// // MIGRATION DRAFT: not included in PLC compilation.
// // Reference: Reference_Project/OPC_Control_FB.scl, object OPC_Control_FB.
// // Types, globals, calls, units and behavior require manual reconciliation.
// // See docs/TIA_Missing_Blocks.md before importing as PLC code.
FUNCTION_BLOCK OPC_Control_FB
// 
//    VAR_INPUT
//       Id : UInt;
//       All_In_Automatic : Bool;
//       VTD_Error : Bool;
//       OPC_Enable : Bool;
//       Clear_OrderTable : Bool;
//    END_VAR
// 
//    VAR_OUTPUT
//       Error_ID : Word;
//    END_VAR
// 
//    VAR
//       Source_Location   : ID_Decoded;
//       Destination_Location   : ID_Decoded;
//       State_Main : UInt;
//       State_VTD : UInt;
//       State_Shuttle : UInt;
//       State_CNV : UInt;
//       T_Wait_Report_Done   : TON;
//    END_VAR
// 
//    VAR_TEMP
//       i : UInt;
//       j : UInt;
//       f : UInt;
//       HMI_Reset : Bool;
//    END_VAR

// // MIGRATION DRAFT: not included in PLC compilation.
// // Reference: Reference_Project/OPC_Control_FB.scl, object OPC_Control_FB.
// // Types, globals, calls, units and behavior require manual reconciliation.
// // See docs/TIA_Missing_Blocks.md before importing as PLC code.
// IF FirstScan THEN
// 	    OPC_Enable := TRUE;
// 	END_IF;
// 
// 	    IF State_CNV > 0 AND State_CNV < 250 THEN
// 
// 	        IF Source_Location.Device_Type = 10 OR Destination_Location.Device_Type = 10 THEN
// 	            IF Control.LCnv_Sys[Id].Cnv_Level[Source_Location.Level].Cnv1.Error
// 	                OR
// 	                Control.LCnv_Sys[Id].Cnv_Level[Destination_Location.Level].Cnv1.Error THEN
// 	                Error_ID.%X3 := TRUE;
// 	                State_CNV := 400;
// 	            END_IF;
// 	        END_IF;
// 
// 	        IF Source_Location.Device_Type = 11 OR Destination_Location.Device_Type = 11 THEN
// 	            IF Control.LCnv_Sys[Id].Cnv_Level[Source_Location.Level].Cnv2.Error
// 	                OR
// 	                Control.LCnv_Sys[Id].Cnv_Level[Destination_Location.Level].Cnv2.Error THEN
// 	                Error_ID.%X3 := TRUE;
// 	                State_CNV := 400;
// 	            END_IF;
// 	        END_IF;
// 
// 	        IF Control.ECnv_Sys[Id].Error THEN
// 	            Error_ID.%X4 := TRUE;
// 	            State_CNV := 400;
// 	        END_IF;
// 	    END_IF;
// 
// 	    IF State_VTD > 0 AND State_VTD < 250 THEN
// 	        IF VTD_Error THEN
// 	            Error_ID.%X5 := TRUE;
// 	            State_VTD := 400;
// 	        END_IF;
// 	    END_IF;
// 
// 	    IF Reset_All THEN
// 	        Error_ID := 0;
// 	    END_IF;
// 
// 	IF State_VTD = 400 OR State_Shuttle = 400 OR State_CNV = 400 THEN
// 	    Error_ID.%X0 := TRUE;
// 	ELSE
// 	    Error_ID.%X0 := FALSE;
// 	    Error_ID.%X6 := FALSE;
// 	    Error_ID.%X7 := FALSE;
// 	    Error_ID.%X8 := FALSE;
// 	END_IF;
// 
// 	IF (Reset_All OR HMI_Reset) AND State_VTD = 400
// 	THEN
// 	    State_VTD := 250;
// 
// 	END_IF;
// 
// 	IF (Reset_All OR HMI_Reset) AND State_Shuttle = 400
// 	THEN
// 	    State_Shuttle := 250;
// 	END_IF;
// 
// 	IF (Reset_All OR HMI_Reset) AND State_CNV = 400
// 	THEN
// 	    State_CNV := 250;
// 	END_IF;
// 
// 	(*
// 	Type of task to be performed:
// 	    1 = Move to Floor
// 	    2 = Shuttle Transfer into VTD
// 	    3 = Shuttle Transfer out of VTD
// 	    4 = Transfer Pallet into VTD
// 	    5 = Transfer Pallet out of VTD
// 	    6 = Transfer Pallet Roller to Roller
// 	    7 = Transfer Pallet Chain to Chain
// 	    8 = Transfer to pick station
// 	    9 = Transfer from Pick station
// 	    10 = Weigh Pallet
// 	    11 = Set chain Cnv as active (lower)
// 	    12 = Set Roller Cnv as active (raise)
// 
// 	    Need to isolate ZZ in XXYYZZ to confirm i = ZZ
// 
// 	    Extract XX (first two digits)
// 	    xx := inputNumber / 10000;
// 
// 	    Extract YY (middle two digits)
// 	    yy := (inputNumber / 100) MOD 100;
// 
// 	    Extract ZZ (last two digits)
// 	    zz := inputNumber MOD 100;
// 	*)
// 
// 
// 	IF All_In_Automatic AND OPC_Enable THEN
// 
// 	        CASE State_Main OF
// 	            0:
// 	                State_Main := 10;
// 
// 	            10:
// 	                IF Control.WCS_OPC_Control[Id].Task_Data_Available AND
// 	                    State_VTD = 0 AND State_Shuttle = 0 AND State_CNV = 0 THEN
// 	                    State_Main := 20;
// 	                END_IF;
// 
// 	            20:
// 	                ID_Decode_F(ID := Control.WCS_OPC_Control[Id].Source_Location,
// 	                              ID_Decoded := Source_Location);
// 	                ID_Decode_F(ID := Control.WCS_OPC_Control[Id].Destination_Location,
// 	                              ID_Decoded := Destination_Location);
// 
// 
// 	                IF Control.WCS_OPC_Control[Id].Task_Type = 1
// 	                    AND NOT Control.VTD[Id].Running THEN
// 	                    State_VTD := 30;
// 	                    Control.WCS_OPC_Control[Id].Task_Data_Available := 0;
// 
// 
// 	                ELSIF Control.WCS_OPC_Control[Id].Task_Type = 2 OR Control.WCS_OPC_Control[Id].Task_Type = 3
// 	                THEN
// 	                    State_Shuttle := 70;
// 	                    Control.WCS_OPC_Control[Id].Task_Data_Available := 0;
// 
// 
// 	                ELSIF (Control.WCS_OPC_Control[Id].Task_Type = 4 OR Control.WCS_OPC_Control[Id].Task_Type = 5)
// 	                THEN
// 	                    State_CNV := 100;
// 	                    Control.WCS_OPC_Control[Id].Task_Data_Available := 0;
// 	                END_IF;
// 	        END_CASE;
// 
// 	            CASE State_VTD OF
// 	                0:
// 	                    ;
// 
// 	                30:
// 	                    State_Main := 0;
// 	                    Control.VTD[Id].Current_Task_Type := INT_TO_UINT(Control.WCS_OPC_Control[Id].Task_Type);
// 	                    Control.VTD[Id].Instruction.Pallet_Type := Control.WCS_OPC_Control[Id].Pallet_Type;
// 	                    Control.VTD[Id].Instruction.Task_ID := INT_TO_UINT(Control.WCS_OPC_Control[Id].Task_ID);
// 	                    Control.VTD[Id].Instruction.Task_Metadata := Control.WCS_OPC_Control[Id].Task_Metadata;
// 	                    Control.VTD[Id].Instruction.Move_To_Level := INT_TO_UINT(Destination_Location.Level);
// 	                    State_VTD := 35;
// 
// 
// 
// 
// 
// 
// 
// 
// 	                35:
// 	                    Control.WCS_OPC_Control[Id].SM_State := Control.VTD[Id].SM_State;
// 	                    IF Control.VTD[Id].Current_Level = Destination_Location.Level THEN
// 
// 	                        Control.WCS_OPC_Control[Id].Movement_Ready := TRUE;
// 	                        State_VTD := 41;
// 	                    ELSIF Control.VTD[Id].Enabled AND Control.VTD[Id].Running THEN
// 	                        Control.WCS_OPC_Control[Id].Movement_Ready := TRUE;
// 	                        State_VTD := 40;
// 	                    END_IF;
// 
// 	                40:
// 	                    Control.WCS_OPC_Control[Id].SM_State := Control.VTD[Id].SM_State;
// 	                    IF Control.VTD[Id].SM_State = 100 THEN
// 	                        State_VTD := 41;
// 	                    END_IF;
// 
// 	                41:
// 	                    T_Wait_Report_Done.TON(IN := TRUE,
// 	                                           PT := T#500ms);
// 	                   IF T_Wait_Report_Done.Q THEN
// 	                       Control.WCS_OPC_Control[Id].Movement_Request_Complete := TRUE;
// 	                       State_VTD := 45;
// 	                   END_IF;
// 
// 	                45:
// 	                    Control.WCS_OPC_Control[Id].SM_State := Control.VTD[Id].SM_State;
// 	                    IF Control.WCS_OPC_Control[Id].Movement_Request_Complete_Ack THEN
// 	                        State_VTD := 250;
// 	                    END_IF;
// 
// 	                250:
// 	                    Control.VTD[Id].Instruction.Reset := FALSE;
// 	                    Control.VTD[Id].Instruction.Pallet_Type := 0;
// 	                    Control.VTD[Id].Instruction.Task_ID := 0;
// 	                    Control.VTD[Id].Instruction.Task_Metadata := '';
// 	                    Control.VTD[Id].Instruction.Move_To_Level := 0;
// 	                    Control.VTD[Id].Current_Task_Type := 0;
// 
// 	                    IF (State_Shuttle = 0 OR State_Shuttle = 250) AND
// 	                        (State_CNV = 0 OR State_CNV = 250) THEN
// 
// 	                        Control.WCS_OPC_Control[Id].SM_State := 0;
// 	                        Control.WCS_OPC_Control[Id].Movement_Ready := FALSE;
// 	                        Control.WCS_OPC_Control[Id].Movement_Request_Complete := FALSE;
// 	                        Control.WCS_OPC_Control[Id].Movement_Request_Complete_Ack := FALSE;
// 	                        Control.WCS_OPC_Control[Id].Pallet_Weight := 0;
// 	                        Control.WCS_OPC_Control[Id].Task_Metadata := '';
// 	                        T_Wait_Report_Done.TON(IN := FALSE,
// 	                                               PT := T#0S);
// 	                       State_VTD := 0;
// 	                    END_IF;
// 
// 	                400:
// 	                    Error_ID.%X6 := TRUE;
// 	                    IF Reset_All OR HMI_Reset
// 	                    THEN
// 	                        Error_ID.%X5 := FALSE;
// 	                        Error_ID.%X6 := FALSE;
// 	                        State_VTD := 250;
// 	                    END_IF;
// 	            END_CASE;
// 	        END_REGION ;
// 
// 	            CASE State_Shuttle OF
// 	                0:
// 	                    ;
// 
// 	                70:
// 	                    State_Main := 0;
// 	                    Control.VTD[Id].Instruction.Task_ID := Control.WCS_OPC_Control[Id].Task_ID;
// 	                    Control.VTD[Id].Instruction.Task_Metadata := Control.WCS_OPC_Control[Id].Task_Metadata;
// 	                    Control.VTD[Id].Instruction.Pallet_Type := Control.WCS_OPC_Control[Id].Pallet_Type;
// 	                    Control.VTD[Id].Current_Task_Type := INT_TO_UINT(Control.WCS_OPC_Control[Id].Task_Type);
// 	                    Control.VTD[Id].Shuttle_Interlock.Shuttle_Interlock_Task_ID := INT_TO_UINT(Control.WCS_OPC_Control[Id].Task_ID);
// 	                    Control.VTD[Id].Shuttle_Interlock.Shuttle_Interlock_Task_Metadata := Control.WCS_OPC_Control[Id].Task_Metadata;
// 	                    Control.VTD[Id].Shuttle_Interlock.Shuttle_ID := INT_TO_UINT(Control.WCS_OPC_Control[Id].Shuttle_ID);
// 	                    Control.VTD[Id].Shuttle_Interlock.Shuttle_Loaded := Control.WCS_OPC_Control[Id].Shuttle_Loaded;
// 	                    Control.VTD[Id].Shuttle_Interlock.Shuttle_Start_Location := Control.WCS_OPC_Control[Id].Source_Location;
// 	                    Control.VTD[Id].Shuttle_Interlock.Shuttle_Target_Location := Control.WCS_OPC_Control[Id].Destination_Location;
// 
// 	                    Control.VTD[Id].Shuttle_Interlock.Interlock_Request := TRUE;
// 	                    State_Shuttle := 75;
// 
// 	                75:
// 	                    Control.WCS_OPC_Control[Id].SM_State := Control.VTD[Id].SM_State;
// 	                    IF Control.VTD[Id].Shuttle_Interlock.Ready_To_Interlock THEN
// 	                        Control.WCS_OPC_Control[Id].Movement_Ready := TRUE;
// 	                        Control.WCS_OPC_Control[Id].Task_Data_Available := FALSE;
// 	                        State_Shuttle := 80;
// 	                    END_IF;
// 
// 	                80:
// 	                    IF Control.VTD[Id].Shuttle_Interlock.Interlock_Complete THEN
// 	                        Control.VTD[Id].Shuttle_Interlock.Interlock_Request := FALSE;
// 	                        Control.WCS_OPC_Control[Id].Movement_Request_Complete := TRUE;
// 	                        State_Shuttle := 90;
// 	                    END_IF;
// 
// 
// 
// 
// 
// 
// 
// 
// 	                90:
// 	                    IF Control.WCS_OPC_Control[Id].Movement_Request_Complete_Ack THEN
// 	                        Control.VTD[Id].Shuttle_Interlock.Interlock_Complete_Ack := TRUE;
// 	                        State_Shuttle := 250;
// 	                    END_IF;
// 
// 	                250:
// 
// 	                    Control.VTD[Id].Shuttle_Interlock.Interlock_Request := FALSE;
// 	                    Control.VTD[Id].Shuttle_Interlock.Shuttle_Start_Location := 0;
// 	                    Control.VTD[Id].Shuttle_Interlock.Shuttle_Target_Location := 0;
// 	                    Control.VTD[Id].Shuttle_Interlock.Shuttle_Loaded := 0;
// 	                    Control.VTD[Id].Shuttle_Interlock.Shuttle_ID := 0;
// 	                    Control.VTD[Id].Shuttle_Interlock.Shuttle_Interlock_Task_ID := 0;
// 	                    Control.VTD[Id].Shuttle_Interlock.Shuttle_Interlock_Task_Metadata := '';
// 	                    Control.VTD[Id].Shuttle_Interlock.Interlock_Complete_Ack := FALSE;
// 
// 	                    IF (State_VTD = 0 OR State_VTD = 250) AND
// 	                        (State_CNV = 0 OR State_CNV = 250) THEN
// 
// 	                        Control.WCS_OPC_Control[Id].SM_State := 0;
// 	                        Control.WCS_OPC_Control[Id].Movement_Ready := FALSE;
// 	                        Control.WCS_OPC_Control[Id].Movement_Request_Complete := FALSE;
// 	                        Control.WCS_OPC_Control[Id].Movement_Request_Complete_Ack := FALSE;
// 	                        Control.WCS_OPC_Control[Id].Task_Metadata := '';
// 	                        T_Wait_Report_Done.TON(IN := FALSE,
// 	                                               PT := T#0S);
// 
// 	                        State_Shuttle := 0;
// 	                    END_IF;
// 
// 	                400:
// 	                    Error_ID.%X7 := TRUE;
// 	                    IF Reset_All OR HMI_Reset
// 	                    THEN
// 	                        Error_ID.%X7 := FALSE;
// 	                        State_Shuttle := 250;
// 	                    END_IF;
// 	            END_CASE;
// 	        END_REGION ;
// 
// 	            CASE State_CNV OF
// 	                0:
// 	                    ;
// 
// 	                100:
// 	                    State_Main := 0;
// 
// 
// 	                    IF Destination_Location.Level >= Settings_DB.VTD[Id].Lowest_Level AND Destination_Location.Level <= Settings_DB.VTD[Id].Highest_Level THEN
// 
// 
// 
// 	                        IF (Destination_Location.Device_Type = 10 AND Control.ECnv_Sys[Id].Cnv_Occupied AND
// 	                            NOT Control.LCnv_Sys[Id].Cnv_Level[Destination_Location.Level].Cnv1.Cnv_Occupied) OR
// 	                            (Destination_Location.Device_Type = 10 AND Destination_Location.Level = 1 AND Source_Location.Device_Type = 0 AND
// 	                            NOT Control.LCnv_Sys[Id].Cnv_Level[Destination_Location.Level].Cnv1.Cnv_Occupied)
// 	                        THEN
// 	                            Control.LCnv_Sys[Id].Cnv_Level[Destination_Location.Level].Cnv1.Instruction.Task_ID := INT_TO_UINT(Control.WCS_OPC_Control[Id].Task_ID);
// 	                            Control.LCnv_Sys[Id].Cnv_Level[Destination_Location.Level].Cnv1.Instruction.Task_Metadata := Control.WCS_OPC_Control[Id].Task_Metadata;
// 	                            Control.LCnv_Sys[Id].Cnv_Level[Destination_Location.Level].Cnv1.Current_Task_Type := INT_TO_UINT(Control.WCS_OPC_Control[Id].Task_Type);
// 	                            Control.LCnv_Sys[Id].Cnv_Level[Destination_Location.Level].Cnv1.Instruction.Transfer_From_ID := Control.WCS_OPC_Control[Id].Source_Location;
// 	                            Control.LCnv_Sys[Id].Cnv_Level[Destination_Location.Level].Cnv1.Instruction.Transfer_To_ID := Control.WCS_OPC_Control[Id].Destination_Location;
// 	                            IF Control.WCS_OPC_Control[Id].Pallet_Type = 'E' AND Control.WCS_OPC_Control[Id].Pallet_Alignment = 'L' THEN
// 	                                Control.LCnv_Sys[Id].Cnv_Level[Destination_Location.Level].Cnv1.Instruction.Pallet_Type := 3;
// 	                            ELSIF Control.WCS_OPC_Control[Id].Pallet_Type = 'E' AND Control.WCS_OPC_Control[Id].Pallet_Alignment = 'R' THEN
// 	                                Control.LCnv_Sys[Id].Cnv_Level[Destination_Location.Level].Cnv1.Instruction.Pallet_Type := 2;
// 	                            END_IF;
// 
// 
// 	                            Control.LCnv_Sys[Id].Cnv_Level[Destination_Location.Level].Cnv1.Instruction.Start_Transfer := TRUE;
// 	                            State_CNV := 105;
// 
// 
// 	                        ELSIF Destination_Location.Device_Type = 11 AND Control.ECnv_Sys[Id].Cnv_Occupied AND
// 	                            NOT Control.LCnv_Sys[Id].Cnv_Level[Destination_Location.Level].Cnv2.Cnv_Occupied
// 	                        THEN
// 	                            Control.LCnv_Sys[Id].Cnv_Level[Destination_Location.Level].Cnv2.Instruction.Task_ID := INT_TO_UINT(Control.WCS_OPC_Control[Id].Task_ID);
// 	                            Control.LCnv_Sys[Id].Cnv_Level[Destination_Location.Level].Cnv2.Instruction.Task_Metadata := Control.WCS_OPC_Control[Id].Task_Metadata;
// 	                            Control.LCnv_Sys[Id].Cnv_Level[Destination_Location.Level].Cnv2.Current_Task_Type := INT_TO_UINT(Control.WCS_OPC_Control[Id].Task_Type);
// 	                            Control.LCnv_Sys[Id].Cnv_Level[Destination_Location.Level].Cnv2.Instruction.Transfer_From_ID := Control.WCS_OPC_Control[Id].Source_Location;
// 	                            Control.LCnv_Sys[Id].Cnv_Level[Destination_Location.Level].Cnv2.Instruction.Transfer_To_ID := Control.WCS_OPC_Control[Id].Destination_Location;
// 	                            IF Control.WCS_OPC_Control[Id].Pallet_Type = 'E' AND Control.WCS_OPC_Control[Id].Pallet_Alignment = 'L' THEN
// 	                                Control.LCnv_Sys[Id].Cnv_Level[Destination_Location.Level].Cnv2.Instruction.Pallet_Type := 3;
// 	                            ELSIF Control.WCS_OPC_Control[Id].Pallet_Type = 'E' AND Control.WCS_OPC_Control[Id].Pallet_Alignment = 'R' THEN
// 	                                Control.LCnv_Sys[Id].Cnv_Level[Destination_Location.Level].Cnv2.Instruction.Pallet_Type := 2;
// 	                            END_IF;
// 
// 
// 	                            Control.LCnv_Sys[Id].Cnv_Level[Destination_Location.Level].Cnv2.Instruction.Start_Transfer := TRUE;
// 	                            State_CNV := 105;
// 
// 
// 	                        ELSIF (Destination_Location.Device_Type = 12 AND Source_Location.Device_Type = 10 AND
// 	                            NOT Control.ECnv_Sys[Id].Cnv_Occupied AND
// 	                            Control.LCnv_Sys[Id].Cnv_Level[Destination_Location.Level].Cnv1.Cnv_Occupied)
// 	                        THEN
// 	                            Control.ECnv_Sys[Id].Instruction.Task_ID := INT_TO_UINT(Control.WCS_OPC_Control[Id].Task_ID);
// 	                            Control.ECnv_Sys[Id].Instruction.Task_Metadata := Control.WCS_OPC_Control[Id].Task_Metadata;
// 	                            Control.ECnv_Sys[Id].Current_Task_Type := INT_TO_UINT(Control.WCS_OPC_Control[Id].Task_Type);
// 	                            Control.ECnv_Sys[Id].Instruction.Transfer_From_ID := Control.WCS_OPC_Control[Id].Source_Location;
// 	                            Control.ECnv_Sys[Id].Instruction.Transfer_To_ID := Control.WCS_OPC_Control[Id].Destination_Location;
// 	                            IF Control.WCS_OPC_Control[Id].Pallet_Type = 'E' AND Control.WCS_OPC_Control[Id].Pallet_Alignment = 'L' THEN
// 	                                Control.ECnv_Sys[Id].Instruction.Pallet_Type := 3;
// 	                            ELSIF Control.WCS_OPC_Control[Id].Pallet_Type = 'E' AND Control.WCS_OPC_Control[Id].Pallet_Alignment = 'R' THEN
// 	                                Control.ECnv_Sys[Id].Instruction.Pallet_Type := 2;
// 	                            ELSIF Control.WCS_OPC_Control[Id].Pallet_Type = 'E' AND Control.WCS_OPC_Control[Id].Pallet_Alignment = 'C' THEN
// 	                                Control.ECnv_Sys[Id].Instruction.Pallet_Type := 4;
// 	                            ELSIF Control.WCS_OPC_Control[Id].Pallet_Type = 'C' THEN
// 	                                Control.ECnv_Sys[Id].Instruction.Pallet_Type := 1;
// 	                            END_IF;
// 
// 
// 	                            Control.ECnv_Sys[Id].Instruction.Start_Transfer := TRUE;
// 	                            State_CNV := 105;
// 
// 
// 	                        ELSIF (Destination_Location.Device_Type = 12 AND Source_Location.Device_Type = 11 AND
// 	                            NOT Control.ECnv_Sys[Id].Cnv_Occupied AND
// 	                            Control.LCnv_Sys[Id].Cnv_Level[Destination_Location.Level].Cnv2.Cnv_Occupied)
// 	                        THEN
// 	                            Control.ECnv_Sys[Id].Instruction.Task_ID := INT_TO_UINT(Control.WCS_OPC_Control[Id].Task_ID);
// 	                            Control.ECnv_Sys[Id].Instruction.Task_Metadata := Control.WCS_OPC_Control[Id].Task_Metadata;
// 	                            Control.ECnv_Sys[Id].Current_Task_Type := INT_TO_UINT(Control.WCS_OPC_Control[Id].Task_Type);
// 	                            Control.ECnv_Sys[Id].Instruction.Transfer_From_ID := Control.WCS_OPC_Control[Id].Source_Location;
// 	                            Control.ECnv_Sys[Id].Instruction.Transfer_To_ID := Control.WCS_OPC_Control[Id].Destination_Location;
// 	                            IF Control.WCS_OPC_Control[Id].Pallet_Type = 'E' AND Control.WCS_OPC_Control[Id].Pallet_Alignment = 'L' THEN
// 	                                Control.ECnv_Sys[Id].Instruction.Pallet_Type := 3;
// 	                            ELSIF Control.WCS_OPC_Control[Id].Pallet_Type = 'E' AND Control.WCS_OPC_Control[Id].Pallet_Alignment = 'R' THEN
// 	                                Control.ECnv_Sys[Id].Instruction.Pallet_Type := 2;
// 	                            ELSIF Control.WCS_OPC_Control[Id].Pallet_Type = 'E' AND Control.WCS_OPC_Control[Id].Pallet_Alignment = 'C' THEN
// 	                                Control.ECnv_Sys[Id].Instruction.Pallet_Type := 4;
// 	                            ELSIF Control.WCS_OPC_Control[Id].Pallet_Type = 'C' THEN
// 	                                Control.ECnv_Sys[Id].Instruction.Pallet_Type := 1;
// 	                            END_IF;
// 
// 
// 	                            Control.ECnv_Sys[Id].Instruction.Start_Transfer := TRUE;
// 	                            State_CNV := 105;
// 
// 
// 	                        ELSIF (Destination_Location.Device_Type = Source_Location.Device_Type AND
// 	                            Control.LCnv_Sys[Id].Cnv_Level[Destination_Location.Level].Cnv1.Cnv_Occupied) AND
// 	                            Control.VTD[Id].Current_Level =  Settings_DB.LCnv_Sys[Id].Cnv_Level[Destination_Location.Level].Cnv1.Cnv_Level
// 	                        THEN
// 	                            Control.LCnv_Sys[Id].Cnv_Level[Destination_Location.Level].Cnv1.Instruction.Task_ID := INT_TO_UINT(Control.WCS_OPC_Control[Id].Task_ID);
// 	                            Control.LCnv_Sys[Id].Cnv_Level[Destination_Location.Level].Cnv1.Instruction.Task_Metadata := Control.WCS_OPC_Control[Id].Task_Metadata;
// 	                            Control.LCnv_Sys[Id].Cnv_Level[Destination_Location.Level].Cnv1.Current_Task_Type := INT_TO_UINT(Control.WCS_OPC_Control[Id].Task_Type);
// 	                            Control.LCnv_Sys[Id].Cnv_Level[Destination_Location.Level].Cnv1.Instruction.Transfer_From_ID := Control.WCS_OPC_Control[Id].Source_Location;
// 	                            Control.LCnv_Sys[Id].Cnv_Level[Destination_Location.Level].Cnv1.Instruction.Transfer_To_ID := Control.WCS_OPC_Control[Id].Destination_Location;
// 	                            IF Control.WCS_OPC_Control[Id].Pallet_Type = 'E' AND Control.WCS_OPC_Control[Id].Pallet_Alignment = 'L' THEN
// 	                                Control.LCnv_Sys[Id].Cnv_Level[Destination_Location.Level].Cnv1.Instruction.Pallet_Type := 3;
// 	                            ELSIF Control.WCS_OPC_Control[Id].Pallet_Type = 'E' AND Control.WCS_OPC_Control[Id].Pallet_Alignment = 'R' THEN
// 	                                Control.LCnv_Sys[Id].Cnv_Level[Destination_Location.Level].Cnv1.Instruction.Pallet_Type := 2;
// 	                            END_IF;
// 
// 
// 	                            Control.LCnv_Sys[Id].Cnv_Level[Destination_Location.Level].Cnv1.Instruction.Pallet_Allignment := TRUE;
// 	                            State_CNV := 112;
// 
// 
// 	                        ELSIF (Destination_Location.Device_Type = Source_Location.Device_Type AND
// 	                            Control.LCnv_Sys[Id].Cnv_Level[Destination_Location.Level].Cnv2.Cnv_Occupied) AND
// 	                            Control.VTD[Id].Current_Level =  Settings_DB.LCnv_Sys[Id].Cnv_Level[Destination_Location.Level].Cnv2.Cnv_Level
// 	                        THEN
// 	                            Control.LCnv_Sys[Id].Cnv_Level[Destination_Location.Level].Cnv2.Instruction.Task_ID := INT_TO_UINT(Control.WCS_OPC_Control[Id].Task_ID);
// 	                            Control.LCnv_Sys[Id].Cnv_Level[Destination_Location.Level].Cnv2.Instruction.Task_Metadata := Control.WCS_OPC_Control[Id].Task_Metadata;
// 	                            Control.LCnv_Sys[Id].Cnv_Level[Destination_Location.Level].Cnv2.Current_Task_Type := INT_TO_UINT(Control.WCS_OPC_Control[Id].Task_Type);
// 	                            Control.LCnv_Sys[Id].Cnv_Level[Destination_Location.Level].Cnv2.Instruction.Transfer_From_ID := Control.WCS_OPC_Control[Id].Source_Location;
// 	                            Control.LCnv_Sys[Id].Cnv_Level[Destination_Location.Level].Cnv2.Instruction.Transfer_To_ID := Control.WCS_OPC_Control[Id].Destination_Location;
// 	                            IF Control.WCS_OPC_Control[Id].Pallet_Type = 'E' AND Control.WCS_OPC_Control[Id].Pallet_Alignment = 'L' THEN
// 	                                Control.LCnv_Sys[Id].Cnv_Level[Destination_Location.Level].Cnv2.Instruction.Pallet_Type := 3;
// 	                            ELSIF Control.WCS_OPC_Control[Id].Pallet_Type = 'E' AND Control.WCS_OPC_Control[Id].Pallet_Alignment = 'R' THEN
// 	                                Control.LCnv_Sys[Id].Cnv_Level[Destination_Location.Level].Cnv2.Instruction.Pallet_Type := 2;
// 	                            END_IF;
// 
// 
// 	                            Control.LCnv_Sys[Id].Cnv_Level[Destination_Location.Level].Cnv2.Instruction.Pallet_Allignment := TRUE;
// 	                            State_CNV := 112;
// 	                        ELSE
// 	                            IF Destination_Location.Device_Type = 10 AND Control.LCnv_Sys[Id].Cnv_Level[Destination_Location.Level].Cnv1.Cnv_Occupied THEN
// 
// 	                                Control.LCnv_Sys[Id].Cnv_Level[Destination_Location.Level].Cnv1.Cnv_Errors.Error_Word_1.%X1 := TRUE;
// 
// 	                            ELSIF Destination_Location.Device_Type = 10 AND Control.LCnv_Sys[Id].Cnv_Level[Destination_Location.Level].Cnv1.Inputs.Shuttle_High THEN
// 
// 	                                Control.LCnv_Sys[Id].Cnv_Level[Destination_Location.Level].Cnv1.Cnv_Errors.Error_Word_1.%X2 := TRUE;
// 
// 	                            ELSIF Destination_Location.Device_Type = 11 AND Control.LCnv_Sys[Id].Cnv_Level[Destination_Location.Level].Cnv2.Cnv_Occupied THEN
// 
// 	                                Control.LCnv_Sys[Id].Cnv_Level[Destination_Location.Level].Cnv2.Cnv_Errors.Error_Word_1.%X1 := TRUE;
// 
// 	                            ELSIF Destination_Location.Device_Type = 11 AND Control.LCnv_Sys[Id].Cnv_Level[Destination_Location.Level].Cnv2.Inputs.Shuttle_High THEN
// 
// 	                                Control.LCnv_Sys[Id].Cnv_Level[Destination_Location.Level].Cnv2.Cnv_Errors.Error_Word_1.%X2 := TRUE;
// 
// 	                            ELSIF Destination_Location.Device_Type = 12 THEN
// 	                                Control.ECnv_Sys[Id].Cnv_Errors.Error_Word_1.%X1 := TRUE;
// 	                            END_IF;
// 
// 	                            State_CNV := 400;
// 	                        END_IF;
// 	                    END_IF;
// 
// 	                105:
// 
// 
// 	                    IF Source_Location.Level >= Settings_DB.VTD[Id].Lowest_Level AND Source_Location.Level <= Settings_DB.VTD[Id].Highest_Level THEN
// 
// 	                        IF Source_Location.Device_Type = 10 AND NOT Control.ECnv_Sys[Id].Cnv_Occupied AND
// 	                            Control.LCnv_Sys[Id].Cnv_Level[Source_Location.Level].Cnv1.Cnv_Occupied
// 	                        THEN
// 	                            Control.LCnv_Sys[Id].Cnv_Level[Source_Location.Level].Cnv1.Instruction.Task_ID := INT_TO_UINT(Control.WCS_OPC_Control[Id].Task_ID);
// 	                            Control.LCnv_Sys[Id].Cnv_Level[Source_Location.Level].Cnv1.Instruction.Task_Metadata := Control.WCS_OPC_Control[Id].Task_Metadata;
// 	                            Control.LCnv_Sys[Id].Cnv_Level[Source_Location.Level].Cnv1.Current_Task_Type := INT_TO_UINT(Control.WCS_OPC_Control[Id].Task_Type);
// 	                            Control.LCnv_Sys[Id].Cnv_Level[Source_Location.Level].Cnv1.Instruction.Transfer_To_ID := Control.WCS_OPC_Control[Id].Destination_Location;
// 	                            Control.LCnv_Sys[Id].Cnv_Level[Source_Location.Level].Cnv1.Instruction.Transfer_From_ID := Control.WCS_OPC_Control[Id].Source_Location;
// 
// 
// 	                            Control.LCnv_Sys[Id].Cnv_Level[Source_Location.Level].Cnv1.Instruction.Start_Transfer := TRUE;
// 	                            State_CNV := 110;
// 
// 
// 	                        ELSIF (Source_Location.Device_Type = 11 AND NOT Control.ECnv_Sys[Id].Cnv_Occupied AND
// 	                            Control.LCnv_Sys[Id].Cnv_Level[Source_Location.Level].Cnv2.Cnv_Occupied) OR
// 	                            (Source_Location.Device_Type = 11 AND Source_Location.Level = 1 AND Destination_Location.Device_Type = 0 AND
// 	                            Control.LCnv_Sys[Id].Cnv_Level[Destination_Location.Level].Cnv2.Cnv_Occupied)
// 	                        THEN
// 	                            Control.LCnv_Sys[Id].Cnv_Level[Source_Location.Level].Cnv2.Instruction.Task_ID := INT_TO_UINT(Control.WCS_OPC_Control[Id].Task_ID);
// 	                            Control.LCnv_Sys[Id].Cnv_Level[Source_Location.Level].Cnv2.Instruction.Task_Metadata := Control.WCS_OPC_Control[Id].Task_Metadata;
// 	                            Control.LCnv_Sys[Id].Cnv_Level[Source_Location.Level].Cnv2.Current_Task_Type := INT_TO_UINT(Control.WCS_OPC_Control[Id].Task_Type);
// 	                            Control.LCnv_Sys[Id].Cnv_Level[Source_Location.Level].Cnv2.Instruction.Transfer_To_ID := Control.WCS_OPC_Control[Id].Destination_Location;
// 	                            Control.LCnv_Sys[Id].Cnv_Level[Source_Location.Level].Cnv2.Instruction.Transfer_From_ID := Control.WCS_OPC_Control[Id].Source_Location;
// 
// 
// 	                            Control.LCnv_Sys[Id].Cnv_Level[Source_Location.Level].Cnv2.Instruction.Start_Transfer := TRUE;
// 	                            State_CNV := 110;
// 
// 
// 	                        ELSIF (Source_Location.Device_Type = 12 AND Destination_Location.Device_Type = 10 AND Control.ECnv_Sys[Id].Cnv_Occupied AND
// 	                            NOT Control.LCnv_Sys[Id].Cnv_Level[Source_Location.Level].Cnv1.Cnv_Occupied)
// 	                        THEN
// 	                            Control.ECnv_Sys[Id].Instruction.Task_ID := INT_TO_UINT(Control.WCS_OPC_Control[Id].Task_ID);
// 	                            Control.ECnv_Sys[Id].Instruction.Task_Metadata := Control.WCS_OPC_Control[Id].Task_Metadata;
// 	                            Control.ECnv_Sys[Id].Current_Task_Type := INT_TO_UINT(Control.WCS_OPC_Control[Id].Task_Type);
// 	                            Control.ECnv_Sys[Id].Instruction.Transfer_To_ID := Control.WCS_OPC_Control[Id].Destination_Location;
// 	                            Control.ECnv_Sys[Id].Instruction.Transfer_From_ID := Control.WCS_OPC_Control[Id].Source_Location;
// 
// 
// 	                            Control.ECnv_Sys[Id].Instruction.Start_Transfer := TRUE;
// 	                            State_CNV := 110;
// 
// 
// 	                        ELSIF (Source_Location.Device_Type = 12 AND Destination_Location.Device_Type = 11 AND Control.ECnv_Sys[Id].Cnv_Occupied AND
// 	                            NOT Control.LCnv_Sys[Id].Cnv_Level[Source_Location.Level].Cnv2.Cnv_Occupied)
// 	                        THEN
// 	                            Control.ECnv_Sys[Id].Instruction.Task_ID := INT_TO_UINT(Control.WCS_OPC_Control[Id].Task_ID);
// 	                            Control.ECnv_Sys[Id].Instruction.Task_Metadata := Control.WCS_OPC_Control[Id].Task_Metadata;
// 	                            Control.ECnv_Sys[Id].Current_Task_Type := INT_TO_UINT(Control.WCS_OPC_Control[Id].Task_Type);
// 	                            Control.ECnv_Sys[Id].Instruction.Transfer_To_ID := Control.WCS_OPC_Control[Id].Destination_Location;
// 	                            Control.ECnv_Sys[Id].Instruction.Transfer_From_ID := Control.WCS_OPC_Control[Id].Source_Location;
// 
// 
// 	                            Control.ECnv_Sys[Id].Instruction.Start_Transfer := TRUE;
// 	                            State_CNV := 110;
// 	                        ELSE
// 	                            State_CNV := 400;
// 	                        END_IF;
// 	                    ELSE
// 	                        State_CNV := 400;
// 	                    END_IF;
// 
// 	                110:
// 	                    Control.WCS_OPC_Control[Id].SM_State := Control.ECnv_Sys[Id].SM_State;
// 
// 	                    IF Control.ECnv_Sys[Id].Enabled AND Control.ECnv_Sys[Id].Running
// 	                    THEN
// 	                        Control.ECnv_Sys[Id].Instruction.Start_Transfer := FALSE;
// 	                        IF (Source_Location.Device_Type = 12 AND Destination_Location.Device_Type = 10) OR
// 	                            (Source_Location.Device_Type = 10 AND Destination_Location.Device_Type = 12) AND
// 	                            Control.LCnv_Sys[Id].Cnv_Level[Control.VTD[Id].Current_Level].Cnv1.Running
// 	                        THEN
// 	                            Control.LCnv_Sys[Id].Cnv_Level[Control.VTD[Id].Current_Level].Cnv1.Instruction.Start_Transfer := FALSE;
// 	                            State_CNV := 115;
// 	                        ELSIF (Source_Location.Device_Type = 12 AND Destination_Location.Device_Type = 11) OR
// 	                            (Source_Location.Device_Type = 11 AND Destination_Location.Device_Type = 12) AND
// 	                            Control.LCnv_Sys[Id].Cnv_Level[Control.VTD[Id].Current_Level].Cnv2.Running
// 	                        THEN
// 	                            Control.LCnv_Sys[Id].Cnv_Level[Control.VTD[Id].Current_Level].Cnv2.Instruction.Start_Transfer := FALSE;
// 	                            State_CNV := 115;
// 	                        END_IF;
// 	                        Control.WCS_OPC_Control[Id].Movement_Ready := TRUE;
// 	                    END_IF;
// 
// 	                112:
// 	                    IF Control.LCnv_Sys[Id].Cnv_Level[Destination_Location.Level].Cnv1.Enabled AND Control.LCnv_Sys[Id].Cnv_Level[Destination_Location.Level].Cnv1.Running
// 	                    THEN
// 	                        Control.WCS_OPC_Control[Id].SM_State := Control.LCnv_Sys[Id].Cnv_Level[Destination_Location.Level].Cnv1.SM_State;
// 	                        Control.LCnv_Sys[Id].Cnv_Level[Destination_Location.Level].Cnv1.Instruction.Pallet_Allignment := FALSE;
// 	                        Control.WCS_OPC_Control[Id].Movement_Ready := TRUE;
// 	                        State_CNV := 116;
// 	                    ELSIF Control.LCnv_Sys[Id].Cnv_Level[Destination_Location.Level].Cnv2.Enabled AND Control.LCnv_Sys[Id].Cnv_Level[Destination_Location.Level].Cnv2.Running
// 	                    THEN
// 	                        Control.WCS_OPC_Control[Id].SM_State := Control.LCnv_Sys[Id].Cnv_Level[Destination_Location.Level].Cnv2.SM_State;
// 	                        Control.LCnv_Sys[Id].Cnv_Level[Destination_Location.Level].Cnv2.Instruction.Pallet_Allignment := FALSE;
// 	                        Control.WCS_OPC_Control[Id].Movement_Ready := TRUE;
// 	                        State_CNV := 116;
// 	                    END_IF;
// 
// 
// 
// 	                115:
// 	                    Control.WCS_OPC_Control[Id].SM_State := Control.ECnv_Sys[Id].SM_State;
// 	                    IF (Source_Location.Device_Type = 12 AND Destination_Location.Device_Type = 10) OR
// 	                        (Source_Location.Device_Type = 10 AND Destination_Location.Device_Type = 12) THEN
// 	                        IF Control.ECnv_Sys[Id].Done AND Control.LCnv_Sys[Id].Cnv_Level[Destination_Location.Level].Cnv1.Done THEN
// 	                            State_CNV := 118;
// 	                        END_IF;
// 	                    ELSIF (Source_Location.Device_Type = 12 AND Destination_Location.Device_Type = 11) OR
// 	                        (Source_Location.Device_Type = 11 AND Destination_Location.Device_Type = 12) THEN
// 	                        IF Control.ECnv_Sys[Id].Done AND Control.LCnv_Sys[Id].Cnv_Level[Destination_Location.Level].Cnv2.Done THEN
// 	                            State_CNV := 118;
// 	                        END_IF;
// 	                    END_IF;
// 
// 	                116:
// 	                        IF Control.LCnv_Sys[Id].Cnv_Level[Destination_Location.Level].Cnv1.Done THEN
// 	                            State_CNV := 118;
// 	                        END_IF;
// 	                        IF Control.LCnv_Sys[Id].Cnv_Level[Destination_Location.Level].Cnv2.Done THEN
// 	                            State_CNV := 118;
// 	                        END_IF;
// 
// 	                118:
// 	                    T_Wait_Report_Done.TON(IN := TRUE,
// 	                                           PT := T#500mS);
// 	                   IF T_Wait_Report_Done.Q THEN
// 	                        Control.WCS_OPC_Control[Id].Movement_Request_Complete := TRUE;
// 	                        State_CNV := 120;
// 	                    END_IF;
// 
// 	                120:
// 	                    Control.WCS_OPC_Control[Id].SM_State := Control.ECnv_Sys[Id].SM_State;
// 	                    IF Control.WCS_OPC_Control[Id].Movement_Request_Complete_Ack THEN
// 	                        State_CNV := 250;
// 	                    END_IF;
// 
// 	                250:
// 	                    Control.ECnv_Sys[Id].Instruction.Reset := FALSE;
// 	                    Control.ECnv_Sys[Id].Instruction.Start_Transfer := FALSE;
// 	                    Control.ECnv_Sys[Id].Instruction.Task_ID := 0;
// 	                    Control.ECnv_Sys[Id].Instruction.Task_Metadata := '';
// 	                    Control.ECnv_Sys[Id].Current_Task_Type := 0;
// 	                    Control.ECnv_Sys[Id].Instruction.Transfer_From_ID := 0;
// 	                    Control.ECnv_Sys[Id].Instruction.Transfer_To_ID := 0;
// 	                    IF Destination_Location.Device_Type = 10 THEN
// 	                        Control.LCnv_Sys[Id].Cnv_Level[Destination_Location.Level].Cnv1.Instruction.Reset := FALSE;
// 	                        Control.LCnv_Sys[Id].Cnv_Level[Destination_Location.Level].Cnv1.Instruction.Start_Transfer := FALSE;
// 	                        Control.LCnv_Sys[Id].Cnv_Level[Destination_Location.Level].Cnv1.Instruction.Task_ID := 0;
// 	                        Control.LCnv_Sys[Id].Cnv_Level[Destination_Location.Level].Cnv1.Instruction.Task_Metadata := '';
// 	                        Control.LCnv_Sys[Id].Cnv_Level[Destination_Location.Level].Cnv1.Current_Task_Type := 0;
// 	                        Control.LCnv_Sys[Id].Cnv_Level[Destination_Location.Level].Cnv1.Instruction.Transfer_From_ID := 0;
// 	                        Control.LCnv_Sys[Id].Cnv_Level[Destination_Location.Level].Cnv1.Instruction.Transfer_To_ID := 0;
// 	                    ELSIF Destination_Location.Device_Type = 11 THEN
// 	                        Control.LCnv_Sys[Id].Cnv_Level[Destination_Location.Level].Cnv2.Instruction.Reset := FALSE;
// 	                        Control.LCnv_Sys[Id].Cnv_Level[Destination_Location.Level].Cnv2.Instruction.Start_Transfer := FALSE;
// 	                        Control.LCnv_Sys[Id].Cnv_Level[Destination_Location.Level].Cnv2.Instruction.Task_ID := 0;
// 	                        Control.LCnv_Sys[Id].Cnv_Level[Destination_Location.Level].Cnv2.Instruction.Task_Metadata := '';
// 	                        Control.LCnv_Sys[Id].Cnv_Level[Destination_Location.Level].Cnv2.Current_Task_Type := 0;
// 	                        Control.LCnv_Sys[Id].Cnv_Level[Destination_Location.Level].Cnv2.Instruction.Transfer_From_ID := 0;
// 	                        Control.LCnv_Sys[Id].Cnv_Level[Destination_Location.Level].Cnv2.Instruction.Transfer_To_ID := 0;
// 	                    ELSIF Source_Location.Device_Type = 10 THEN
// 	                        Control.LCnv_Sys[Id].Cnv_Level[Source_Location.Level].Cnv1.Instruction.Reset := FALSE;
// 	                        Control.LCnv_Sys[Id].Cnv_Level[Source_Location.Level].Cnv1.Instruction.Start_Transfer := FALSE;
// 	                        Control.LCnv_Sys[Id].Cnv_Level[Source_Location.Level].Cnv1.Instruction.Task_ID := 0;
// 	                        Control.LCnv_Sys[Id].Cnv_Level[Source_Location.Level].Cnv1.Instruction.Task_Metadata := '';
// 	                        Control.LCnv_Sys[Id].Cnv_Level[Source_Location.Level].Cnv1.Current_Task_Type := 0;
// 	                        Control.LCnv_Sys[Id].Cnv_Level[Source_Location.Level].Cnv1.Instruction.Transfer_From_ID := 0;
// 	                        Control.LCnv_Sys[Id].Cnv_Level[Source_Location.Level].Cnv1.Instruction.Transfer_To_ID := 0;
// 	                    ELSIF Destination_Location.Device_Type = 11 THEN
// 	                        Control.LCnv_Sys[Id].Cnv_Level[Source_Location.Level].Cnv2.Instruction.Reset := FALSE;
// 	                        Control.LCnv_Sys[Id].Cnv_Level[Source_Location.Level].Cnv2.Instruction.Start_Transfer := FALSE;
// 	                        Control.LCnv_Sys[Id].Cnv_Level[Source_Location.Level].Cnv2.Instruction.Task_ID := 0;
// 	                        Control.LCnv_Sys[Id].Cnv_Level[Source_Location.Level].Cnv2.Instruction.Task_Metadata := '';
// 	                        Control.LCnv_Sys[Id].Cnv_Level[Source_Location.Level].Cnv2.Current_Task_Type := 0;
// 	                        Control.LCnv_Sys[Id].Cnv_Level[Source_Location.Level].Cnv2.Instruction.Transfer_From_ID := 0;
// 	                        Control.LCnv_Sys[Id].Cnv_Level[Source_Location.Level].Cnv2.Instruction.Transfer_To_ID := 0;
// 	                    END_IF;
// 
// 
// 
// 
// 	                        Control.WCS_OPC_Control[Id].SM_State := 0;
// 	                        Control.WCS_OPC_Control[Id].Movement_Ready := FALSE;
// 	                        Control.WCS_OPC_Control[Id].Movement_Request_Complete := FALSE;
// 	                        Control.WCS_OPC_Control[Id].Movement_Request_Complete_Ack := FALSE;
// 	                        Control.WCS_OPC_Control[Id].Task_Metadata := '';
// 	                        T_Wait_Report_Done.TON(IN := FALSE,
// 	                                               PT := T#0S);
// 
// 	                        State_CNV := 0;
// 
// 
// 	                    400:
// 	                        Error_ID.%X8 := TRUE;
// 	                        IF Reset_All OR HMI_Reset THEN
// 	                            Error_ID.%X3 := FALSE;
// 	                            Error_ID.%X4 := FALSE;
// 	                            Error_ID.%X8 := FALSE;
// 	                            State_CNV := 250;
// 	                    END_IF;
// 	            END_CASE;
// 	        END_REGION ;
// 
// 	ELSIF All_In_Automatic AND NOT OPC_Enable THEN
// 
// 
// 
// 	    Control.WCS_OPC_Control[Id].SM_State := 0;
// 	    Control.WCS_OPC_Control[Id].Movement_Ready := FALSE;
// 	    Control.WCS_OPC_Control[Id].Movement_Request_Complete := FALSE;
// 
// 
// 	    Control.WCS_OPC_Control[Id].Task_Type := 0;
// 	    Control.WCS_OPC_Control[Id].Pallet_Type := 'C';
// 	    Control.WCS_OPC_Control[Id].Task_ID := 0;
// 	    Control.WCS_OPC_Control[Id].Task_Metadata := '';
// 	    Control.WCS_OPC_Control[Id].Source_Location := 0;
// 	    Control.WCS_OPC_Control[Id].Destination_Location := 0;
// 	    Destination_Location.Level := 0;
// 	    Source_Location.Level := 0;
// 	    Control.WCS_OPC_Control[Id].Shuttle_ID := 0;
// 	    Control.WCS_OPC_Control[Id].Shuttle_Loaded := FALSE;
// 
// 
// 	    Control.VTD[Id].Instruction.Reset := FALSE;
// 	    Control.VTD[Id].Instruction.Pallet_Type := 0;
// 	    Control.VTD[Id].Instruction.Task_ID := 0;
// 	    Control.VTD[Id].Instruction.Task_Metadata := '';
// 	    Control.ECnv_Sys[Id].Current_Task_Type := 0;
// 	    Control.VTD[Id].Instruction.Move_To_Level := 99;
// 	    Control.VTD[Id].Current_Task_Type := 0;
// 
// 
// 	    Control.VTD[Id].Shuttle_Interlock.Interlock_Request := FALSE;
// 	    Control.VTD[Id].Shuttle_Interlock.Shuttle_Start_Location := 0;
// 	    Control.VTD[Id].Shuttle_Interlock.Shuttle_Target_Location := 0;
// 	    Control.VTD[Id].Shuttle_Interlock.Shuttle_Loaded := 0;
// 	    Control.VTD[Id].Shuttle_Interlock.Shuttle_ID := 0;
// 	    Control.VTD[Id].Shuttle_Interlock.Shuttle_Interlock_Task_ID := 0;
// 	    Control.VTD[Id].Shuttle_Interlock.Shuttle_Interlock_Task_Metadata := '';
// 
// 
// 	    Control.ECnv_Sys[Id].Instruction.Reset := FALSE;
// 
// 	    Control.ECnv_Sys[Id].Instruction.Start_Transfer := FALSE;
// 	    Control.ECnv_Sys[Id].Instruction.Task_ID := 0;
// 	    Control.ECnv_Sys[Id].Instruction.Task_Metadata := '';
// 	    Control.ECnv_Sys[Id].Instruction.Transfer_From_ID := 0;
// 	    Control.ECnv_Sys[Id].Instruction.Transfer_To_ID := 0;
// 
// 	    FOR i := Settings_DB.VTD[Id].Lowest_Level TO Settings_DB.VTD[Id].Highest_Level DO
// 	        Control.LCnv_Sys[Id].Cnv_Level[i].Cnv1.Instruction.Reset := FALSE;
// 	        Control.LCnv_Sys[Id].Cnv_Level[i].Cnv1.Instruction.Start_Transfer := FALSE;
// 	        Control.LCnv_Sys[Id].Cnv_Level[i].Cnv1.Instruction.Task_ID := 0;
// 	        Control.LCnv_Sys[Id].Cnv_Level[i].Cnv1.Instruction.Task_Metadata := '';
// 	        Control.LCnv_Sys[Id].Cnv_Level[i].Cnv1.Current_Task_Type := 0;
// 	        Control.LCnv_Sys[Id].Cnv_Level[i].Cnv1.Instruction.Transfer_From_ID := 0;
// 	        Control.LCnv_Sys[Id].Cnv_Level[i].Cnv1.Instruction.Transfer_To_ID := 0;
// 
// 	        Control.LCnv_Sys[Id].Cnv_Level[i].Cnv2.Instruction.Reset := FALSE;
// 	        Control.LCnv_Sys[Id].Cnv_Level[i].Cnv2.Instruction.Start_Transfer := FALSE;
// 	        Control.LCnv_Sys[Id].Cnv_Level[i].Cnv2.Instruction.Task_ID := 0;
// 	        Control.LCnv_Sys[Id].Cnv_Level[i].Cnv2.Instruction.Task_Metadata := '';
// 	        Control.LCnv_Sys[Id].Cnv_Level[i].Cnv2.Current_Task_Type := 0;
// 	        Control.LCnv_Sys[Id].Cnv_Level[i].Cnv2.Instruction.Transfer_From_ID := 0;
// 	        Control.LCnv_Sys[Id].Cnv_Level[i].Cnv2.Instruction.Transfer_To_ID := 0;
// 	    END_FOR;
// 	END_IF;
// 
// 	    IF Clear_OrderTable THEN
// 	        State_Main := 0;
// 	        State_VTD := 250;
// 	        State_Shuttle := 250;
// 	        State_CNV := 250;
// 	        Control.WCS_OPC_Control[Id].Task_Data_Available := 0;
// 	    END_IF;
// 
// 
// 	    FOR f := 1 TO Settings_DB.System.Shuttle_Count DO
// 	        Control.Shuttles_Position[f].x := Shuttle_MQTT_DB.Shuttle_MQTT[f].Message.Shuttle_Status.Position_X;
// 	        Control.Shuttles_Position[f].y := Shuttle_MQTT_DB.Shuttle_MQTT[f].Message.Shuttle_Status.Position_Y;
// 	    END_FOR;
// 
// 
// 
// 	HMI_Reset := (Screen_DB_1.Reset_All[1] AND
// 	(HMI_Box_Connected_1 = 1) OR (HMI_Box_Connected_1 = 2) OR (HMI_Box_Connected_1 = 3) OR (HMI_Box_Connected_1 = 4) OR (HMI_Box_Connected_1 = 5) OR
// 	(HMI_Box_Connected_1 = 11 AND KEY_REMOTE_LOCAL_L1___CH1_1_) OR
// 	(HMI_Box_Connected_1 = 12 AND KEY_REMOTE_LOCAL_L2___CH1_1_) OR
// 	(HMI_Box_Connected_1 = 13 AND KEY_REMOTE_LOCAL_L3___CH1_1_) OR
// 	(HMI_Box_Connected_1 = 14 AND KEY_REMOTE_LOCAL_L4___CH1_1_) OR
// 	(HMI_Box_Connected_1 = 15 AND KEY_REMOTE_LOCAL_L5___CH1_1_) OR
// 	(HMI_Box_Connected_1 = 16 AND KEY_REMOTE_LOCAL_L6___CH1_1_) OR
// 	(HMI_Box_Connected_1 = 17 AND KEY_REMOTE_LOCAL_L7___CH1_1_) OR
// 	(HMI_Box_Connected_1 = 18 AND KEY_REMOTE_LOCAL_L8___CH1_1_) OR
// 	(HMI_Box_Connected_1 = 21 AND KEY_REMOTE_LOCAL_L1___CH1_2_) OR
// 	(HMI_Box_Connected_1 = 22 AND KEY_REMOTE_LOCAL_L2___CH1_2_) OR
// 	(HMI_Box_Connected_1 = 23 AND KEY_REMOTE_LOCAL_L3___CH1_2_) OR
// 	(HMI_Box_Connected_1 = 24 AND KEY_REMOTE_LOCAL_L4___CH1_2_) OR
// 	(HMI_Box_Connected_1 = 25 AND KEY_REMOTE_LOCAL_L5___CH1_2_) OR
// 	(HMI_Box_Connected_1 = 26 AND KEY_REMOTE_LOCAL_L6___CH1_2_) OR
// 	(HMI_Box_Connected_1 = 27 AND KEY_REMOTE_LOCAL_L7___CH1_2_) OR
// 	(HMI_Box_Connected_1 = 28 AND KEY_REMOTE_LOCAL_L8___CH1_2_) OR
// 	(HMI_Box_Connected_1 = 31 AND KEY_REMOTE_LOCAL_L1___CH1_3_) OR
// 	(HMI_Box_Connected_1 = 32 AND KEY_REMOTE_LOCAL_L2___CH1_3_) OR
// 	(HMI_Box_Connected_1 = 33 AND KEY_REMOTE_LOCAL_L3___CH1_3_) OR
// 	(HMI_Box_Connected_1 = 34 AND KEY_REMOTE_LOCAL_L4___CH1_3_) OR
// 	(HMI_Box_Connected_1 = 35 AND KEY_REMOTE_LOCAL_L5___CH1_3_) OR
// 	(HMI_Box_Connected_1 = 36 AND KEY_REMOTE_LOCAL_L6___CH1_3_) OR
// 	(HMI_Box_Connected_1 = 37 AND KEY_REMOTE_LOCAL_L7___CH1_3_) OR
// 	(HMI_Box_Connected_1 = 38 AND KEY_REMOTE_LOCAL_L8___CH1_3_) OR
// 	(HMI_Box_Connected_1 = 41 AND KEY_REMOTE_LOCAL_L1___CH1_4_) OR
// 	(HMI_Box_Connected_1 = 42 AND KEY_REMOTE_LOCAL_L2___CH1_4_) OR
// 	(HMI_Box_Connected_1 = 43 AND KEY_REMOTE_LOCAL_L3___CH1_4_) OR
// 	(HMI_Box_Connected_1 = 44 AND KEY_REMOTE_LOCAL_L4___CH1_4_) OR
// 	(HMI_Box_Connected_1 = 45 AND KEY_REMOTE_LOCAL_L5___CH1_4_) OR
// 	(HMI_Box_Connected_1 = 46 AND KEY_REMOTE_LOCAL_L6___CH1_4_) OR
// 	(HMI_Box_Connected_1 = 47 AND KEY_REMOTE_LOCAL_L7___CH1_4_) OR
// 	(HMI_Box_Connected_1 = 48 AND KEY_REMOTE_LOCAL_L8___CH1_4_) OR
// 	(HMI_Box_Connected_1 = 51 AND KEY_REMOTE_LOCAL_L1___CH1_5_) OR
// 	(HMI_Box_Connected_1 = 52 AND KEY_REMOTE_LOCAL_L2___CH1_5_) OR
// 	(HMI_Box_Connected_1 = 53 AND KEY_REMOTE_LOCAL_L3___CH1_5_) OR
// 	(HMI_Box_Connected_1 = 54 AND KEY_REMOTE_LOCAL_L4___CH1_5_) OR
// 	(HMI_Box_Connected_1 = 55 AND KEY_REMOTE_LOCAL_L5___CH1_5_) OR
// 	(HMI_Box_Connected_1 = 56 AND KEY_REMOTE_LOCAL_L6___CH1_5_) OR
// 	(HMI_Box_Connected_1 = 57 AND KEY_REMOTE_LOCAL_L7___CH1_5_) OR
// 	(HMI_Box_Connected_1 = 58 AND KEY_REMOTE_LOCAL_L8___CH1_5_));

END_FUNCTION_BLOCK

(* stored: Version 1.1.0.1
   POU OPC_Control_FB: Id {4b22b142-7a62-51de-b74c-3fbf01b234a1}, SpecialFunc None *)
